(*
SPDX-FileCopyrightText: c 2026 Oleksandr Tiutyk <trofimich@gmail.com>
SPDX-License-Identifier: MIT
License: https://opensource.org/license/mit
*)

(*!
<summary>Checks full and windowed joining and cursor reuse after insufficient capacity.</summary>
<description>
Uses one task and stays at a stable address while assertions are bound to this instance.
</description>
*)

{attribute 'no_assign'}
{attribute 'no_explicit_call' := 'do not call this function block directly'}
FUNCTION_BLOCK StringJoinTest EXTENDS TOF_Testing.SingleCycleTest
VAR_STAT
	{attribute 'hide'}
	_ClassName : STRING := __POUNAME();
END_VAR
VAR
	_Source : STRING := '123 , , 456, 789 ,0';
	_Splitter : TOF_Core.StringSplittingEnumerator;
END_VAR

(*!
<summary>Checks full and windowed joining and cursor reuse after insufficient capacity.</summary>
<description>
Owns a persistent cursor and its borrowed source. Reset releases the current fragment before the result is reported.
</description>
*)
METHOD PROTECTED ExecuteTest
VAR
	separator : STRING := ',';
	joined : STRING := 'old target';
	shortTarget : STRING(2);
	accepted : BOOL;
END_VAR
_Splitter := TOF_Core.Strings.CreateSplitter(sourceString := _Source, separator := separator);
TOF_Core.Strings.Join(targetString := joined, separator := separator, sourceEnumerator := _Splitter);
Assert.ThatBool(
	actual := joined = _Source,
	message := "Unrestricted Join must reconstruct all fragments including their whitespace"
).IsTrue();

_Splitter.Reset();
_Splitter := TOF_Core.Strings.CreateSplitter(
	sourceString := _Source,
	separator := separator,
	maxCount := 3,
	trimEntries := TRUE,
	removeEmptyEntries := TRUE
);
TOF_Core.Strings.Join(
	targetString := joined,
	separator := separator,
	sourceEnumerator := _Splitter,
	startIndex := 1,
	count := 2
);
Assert.ThatBool(
	actual := joined = '456,789',
	message := "The requested window must contain fragments 1 and 2"
).IsTrue();

_Splitter.Reset();
accepted := TOF_Core.Strings.TryJoin(targetString := shortTarget, separator := separator, sourceEnumerator := _Splitter);
Assert.ThatBool(
	actual := accepted,
	message := "TryJoin must reject a target too small for the first fragment"
).IsFalse();

_Splitter.Reset();
accepted := TOF_Core.Strings.TryJoin(
	targetString := joined,
	separator := separator,
	sourceEnumerator := _Splitter,
	count := 1
);
Assert.ThatBool(
	actual := accepted AND_THEN joined = '123',
	message := "After Reset, TryJoin must restart and replace the old target text"
).IsTrue();
END_METHOD

(*!
<summary>Resets the splitter and releases any active fragment before reporting.</summary>
<description>
Safe after partial initialization and after explicit cleanup in the scenario.
</description>
*)
METHOD PROTECTED AfterTest
_Splitter.Reset();
END_METHOD

//! <summary>Borrows the concrete class name. Callers must not modify it.</summary>
{attribute 'monitoring' := 'call'}
PROPERTY ClassName : REFERENCE TO STRING
GET
ClassName REF= _ClassName;
END_GET
END_PROPERTY

//! <summary>Borrows the compiler-initialized namespace name. Callers must not modify it.</summary>
{attribute 'monitoring' := 'call'}
PROPERTY NamespaceName : REFERENCE TO STRING
GET
NamespaceName REF= CurrentNamespace.Name;
END_GET
END_PROPERTY

//! <summary>Reports the concrete instance size in bytes.</summary>
{attribute 'monitoring' := 'call'}
PROPERTY SelfSize : ULINT
GET
SelfSize := XSIZEOF(THIS^);
END_GET
END_PROPERTY

END_FUNCTION_BLOCK

(* stored: Version 1.1.0.1
   POU StringJoinTest: Id {c8768789-bd41-4bd0-b0ca-488801c6d010}, SpecialFunc None
   Method ExecuteTest: Id {54c50b31-ade0-4d37-9420-f9ab6f4b0f3c}
   Method AfterTest: Id {43a92498-5d4d-41dd-8275-2820bc42fa64}
   Property ClassName: Id {79e0b534-a61f-4f38-9fe8-0da2851208ba}
   Get Get: Id {215a8ae3-1ea4-4b91-bc49-8cc0d4dee3ec}
   Property NamespaceName: Id {cac03636-e2ff-40d5-9305-c95241594bce}
   Get Get: Id {d6ad1ed0-55ec-4946-8516-f34873e5f8ad}
   Property SelfSize: Id {732342f9-774b-46a2-ac81-3f2605faa1b4}
   Get Get: Id {4becf984-735f-4f34-aee9-d17a1a5c3596} *)
